// TIA Portal V21 export
DATA_BLOCK "IDB_AnaGlobalAccess"   // DB11
// stored: InstanceOfName FB_AnaGlobalAccess, InstanceOfType FB
"FB_AnaGlobalAccess"
   // VAR_OUTPUT
   //    Speed : Real;
   // END_VAR
BEGIN
END_DATA_BLOCK
